TYPE ST_PolarIIChamber_NozzlePortServiceCtrl :
STRUCT
	Nozzle : ARRAY[1..3] OF ST_PolarIIChamber_PortNozzleSupplyServiceCtrl;
	DrainSelect1 : ST_ServiceCtrl;
	DrainSelect2 : ST_ServiceCtrl;
	DrainSelect3 : ST_ServiceCtrl;
END_STRUCT
END_TYPE

(* stored: Version 1.1.0.1, ProductVersion 3.1.4026.18
   DUT ST_PolarIIChamber_NozzlePortServiceCtrl: Id {14000000-0000-0000-0000-000000000055} *)
